// TIA Portal V20 export
Screen "01_ScreenLayout"  1366x768
  ScreenItem "swHeader" at 0,1 size 1366x65  Type=HmiScreenWindow
  ScreenItem "swAlarm" at 0,65 size 1276x30  Type=HmiScreenWindow
  ScreenItem "swMainSmall" at 1276,65 size 90x703  Type=HmiScreenWindow
  ScreenItem "swContent" at 0,95 size 1276x673  Type=HmiScreenWindow
